// TIA Portal V15.1 export
DATA_BLOCK "HmiAlm"   // DB6
{ S7_Optimized_Access := 'TRUE' }
VERSION : 0.1
// stored: AutoNumber false, MemoryReserve 100
   VAR
      Common : Word;   // 0007 / H-05: x0 E-STOP active or not reset [C01]; x1 Scrubber trip: high pressure PSH-101 [C03 / C06a (PH proposal: cause memory)]; x2 Scrubber trip: high-high level LSHH-103 [C05 / C06a (PH proposal: cause memory)]; x3 Scrubber held after power-up: RESET required [S-01 / C06a (PH proposal)]; x4 Scrubber high level LSH-102 [C04 (Client)]; x5 Setting rejected: out of range [R-11]; x6 Scrubber drain open too long: drain closed [C04a]; x7 LSH-102 fault: LSHH-103 without LSH-102 [C04b]
      BR01 : Word;   // 0007 / H-05: x0 BR01 stopped by E-STOP: RESET + START [C01]; x1 BR01 thermocouple fault [C07d]; x2 BR01 burner lockout [C07e]; x3 BR01 failed to start [C07f]; x4 BR01 stopped by itself [C07g]; x5 BR01 RUN without request [R-09]; x6 TK01 level low: burner held [C07a (PH proposal: alarm; Client: permissive)]
      BR02 : Word;   // 0007 / H-05: x0 BR02 stopped by E-STOP: RESET + START [C01]; x1 BR02 thermocouple fault [C08d]; x2 BR02 burner lockout [C08e]; x3 BR02 failed to start [C08f]; x4 BR02 stopped by itself [C08g]; x5 BR02 RUN without request [R-09]; x6 TK02 level low: burner held [C08a (PH proposal: alarm; Client: permissive)]
   END_VAR
BEGIN
END_DATA_BLOCK
